Staubli VAL3: progTemp.dtx

public progItem pProgItem{}
  [Key1]
    progTemplate pProgTemplate
      [0]
        forItem fForItem
          [0]
            bool bIOdisable
            num nLoopValue
            string sForTRAJ
            string sIOindex
        ifItem iIfItem
          [0]
            bool bANDOR[2]
            num nSigIndex[3]
            num nSigType[3]
            num nValue[3]
        num nType
        switchItem sSwitchItem
          [0]
            bool bIOdisable
            num nSwitchValue
            string sIOValue
        string sTRAJname
